Fanuc KAREL source: kf00054.KL

-- PROVISIONAL review KL for V1013-1; original PC SHA256 6abe4517b66a4608bee078a133812307e0a8ebe5f482341c8cc15917644d6cf5
-- Incomplete behavior may be omitted. Consult companion uncertainty JSON. Do not deploy.
PROGRAM KF00054
%NOLOCKGROUP
VAR
  I : INTEGER
  J : INTEGER
  X : REAL
  Y : REAL
  B : BOOLEAN
  C : BOOLEAN
  TXT : STRING[80]
  TXT2 : STRING[80]
  STATUS : INTEGER
-- UNRESOLVED_DECL AI type=002010
-- UNRESOLVED_DECL BI type=002010
-- UNRESOLVED_DECL P type=000102
-- UNRESOLVED_DECL JP type=000199
-- UNRESOLVED_DECL PF type=000101
-- UNRESOLVED_DECL V1 type=000013
-- UNRESOLVED_DECL V2 type=000013
BEGIN
  -- UNRESOLVED_PC offsets 5-12; opcodes 9D,23
  -- UNRESOLVED_PC offsets 17-22; opcodes 7A
  -- UNRESOLVED_PC offsets 27-38; opcodes 2E,23
  -- UNRESOLVED_PC offsets 43-54; opcodes 2E,23
  -- UNRESOLVED_PC offsets 59-63; opcodes 7F
END KF00054
